// TIA Portal V20 export
FUNCTION_BLOCK "PR_HIPOTTestSeq_Soft2.0 1_workflow_cd2a65"   // FB45, LAD
{ S7_Optimized_Access := 'TRUE' }
// stored: MemoryReserve 100, SetENOAutomatically false
   VAR_INPUT
      iAutoRunning : Bool;
      iFaultReset : Bool;
      iHiPotProbeUp : Bool;
      iHiPotTestOver : Bool;
      iHiPotTestProbeDown : Bool;
      iPartPresent : Bool;
      iPressProbeUp : Bool;
      iReset_fault : Bool;
      iShuttleAtHiPotTest : Bool;
      iSstMode : Bool;
      iSstPB : Bool;
      iStartFrmShuttleSeq : Bool;
      iTestProbeDown : Bool;
      iTestProbeUp : Bool;
      iTestProbesUp : Bool;
      iThicknessTestOver : Bool;
      iScanOK : Bool;
      iScanNOK : Bool;
      iRetryCount : Int;
      iForcedAccept : Bool;
      iRetry : Bool;
   END_VAR
   VAR_OUTPUT
      qHiPotTestOver : Bool;
      qStateNo : Int;
      qMessage : Array[0..2] of Bool;
   END_VAR
   VAR
      c20_ChkRecoveryStatus_T1 : Bool;
      c20_ChkRecoveryStatus_T2 : Bool;
      c20_ChkRecoveryStatus_T3 : Bool;
      c20_ChkRecoveryStatus_T4 : Bool;
      c50_ChkPartPresentShuttlePos_T1 : Bool;
      c50_ChkPartPresentShuttlePos_T2 : Bool;
      s100_WtHiPotTestProbesDown : Bool;
      s100_WtHiPotTestProbesDown_T1 : Bool;
      s10_WtStartFrmShuttleSeq : Bool;
      s10_WtStartFrmShuttleSeq_T1 : Bool;
      s110_WtHiPotTestOver : Bool;
      s110_WtHiPotTestOver_T1 : Bool;
      s120_WtHiPotProbeUp : Bool;
      s120_WtHiPotProbeUp_T1 : Bool;
      s130_WtPressProbesUp : Bool;
      s130_WtPressProbesUp_T1 : Bool;
      s140_WtStartLow : Bool;
      s140_WtStartLow_T1 : Bool;
      s1_WtResetRel : Bool;
      s1_WtResetRel_T1 : Bool;
      s20_ChkRecoveryStatus : Bool;
      s20_ChkRecoveryStatus_T1 : Bool;
      s20_ChkRecoveryStatus_T2 : Bool;
      s20_ChkRecoveryStatus_T3 : Bool;
      s20_ChkRecoveryStatus_T4 : Bool;
      s30_WtOperatorAck : Bool;
      s30_WtOperatorAck_T1 : Bool;
      s40_WtAllSlidesHome : Bool;
      s40_WtAllSlidesHome_T1 : Bool;
      s50_ChkPartPresentShuttlePos : Bool;
      s50_ChkPartPresentShuttlePos_T1 : Bool;
      s50_ChkPartPresentShuttlePos_T2 : Bool;
      s75_WtScanOver : Bool;
      s75_WtScanOver_T1 : Bool;
      s75_WtScanOver_T2 : Bool;
      s76_ChkReryCountOver : Bool;
      s76_ChkRetryCountOver_T1 : Bool;
      s76_ChkRetryCountOver_T2 : Bool;
      s77_WtOperatorDecision : Bool;
      s77_WtOperatorDecision_T1 : Bool;
      s77_WtOperatorDecision_T2 : Bool;
      s70_WtPartPresentShuttlePos : Bool;
      s70_WtPartPresentShuttlePos_T1 : Bool;
      s80_WtTestProbeDown : Bool;
      s80_WtTestProbeDown_T1 : Bool;
      s90_WtThicknessTestOver : Bool;
      s90_WtThicknessTestOver_T1 : Bool;
      sAbnormalStatus : Bool;
      sHiPotTestInProgress : Bool;
      sSst : Bool;
      sSstPulse : Bool;
      sSstRise : Bool;
      sStWtResetRel : Bool;
      sStWtResetRel_T1 : Bool;
      sThicknessTestInProgress : Bool;
      sScanRetryCount : Int;
   END_VAR
   VAR_TEMP
      tOne : Bool;
   END_VAR
   VAR_TEMP   // added for the SCL form of the ladder/FBD networks
      _w1 : Bool;
      _w2 : Bool;
      _w3 : Bool;
   END_VAR
BEGIN

REGION Network 1
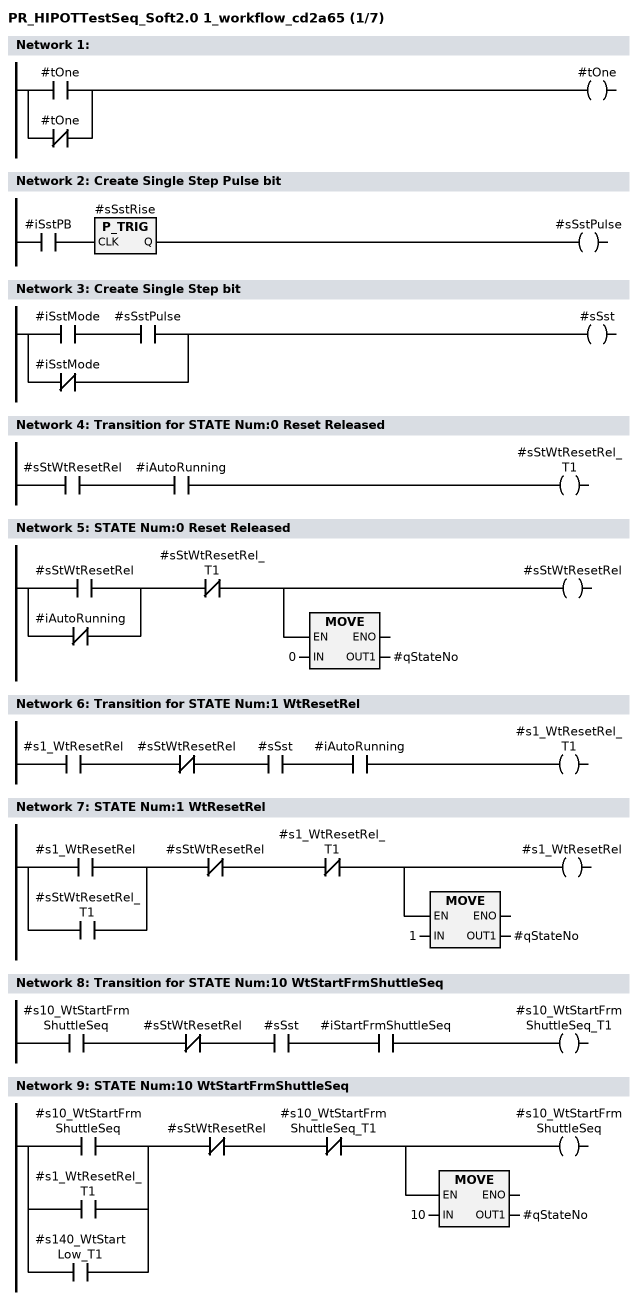
   RUNG wire#powerrail
      Contact( #tOne )
      wire#w1
      Coil( #tOne )
   END_RUNG
   RUNG wire#powerrail
      I_Contact( #tOne )
   END_RUNG wire#w1
   // the same network as SCL:
   #tOne := #tOne OR NOT #tOne;
END_REGION

REGION Network 2: Create Single Step Pulse bit
   RUNG wire#powerrail
      Contact( #iSstPB )
      P_Trig( #sSstRise )
      Coil( #sSstPulse )
   END_RUNG
   // the same network as SCL:
   #_w1 := #iSstPB AND NOT #sSstRise;   // rising edge
   #sSstRise := #iSstPB;
   #sSstPulse := #_w1;
END_REGION

REGION Network 3: Create Single Step bit
   RUNG wire#powerrail
      Contact( #iSstMode )
      Contact( #sSstPulse )
      wire#w1
      Coil( #sSst )
   END_RUNG
   RUNG wire#powerrail
      I_Contact( #iSstMode )
   END_RUNG wire#w1
   // the same network as SCL:
   #sSst := (#iSstMode AND #sSstPulse) OR NOT #iSstMode;
END_REGION

REGION Network 4: Transition for STATE Num:0 Reset Released
   RUNG wire#powerrail
      Contact( #sStWtResetRel )
      Contact( #iAutoRunning )
      Coil( #sStWtResetRel_T1 )
   END_RUNG
   // the same network as SCL:
   #sStWtResetRel_T1 := #sStWtResetRel AND #iAutoRunning;
END_REGION

REGION Network 5: STATE Num:0 Reset Released
   RUNG wire#powerrail
      Contact( #sStWtResetRel )
      wire#w1
      I_Contact( #sStWtResetRel_T1 )
      wire#w2
      Coil( #sStWtResetRel )
   END_RUNG
   RUNG wire#powerrail
      I_Contact( #iAutoRunning )
   END_RUNG wire#w1
   RUNG wire#w2
      { S7_GenerateENO := "TRUE" } Move(in := 0, out1 => #qStateNo)
   END_RUNG
   // the same network as SCL:
   #sStWtResetRel := (#sStWtResetRel OR NOT #iAutoRunning) AND NOT #sStWtResetRel_T1;
   IF #sStWtResetRel THEN #qStateNo := 0; END_IF;
END_REGION

REGION Network 6: Transition for STATE Num:1 WtResetRel
   RUNG wire#powerrail
      Contact( #s1_WtResetRel )
      I_Contact( #sStWtResetRel )
      Contact( #sSst )
      Contact( #iAutoRunning )
      Coil( #s1_WtResetRel_T1 )
   END_RUNG
   // the same network as SCL:
   #s1_WtResetRel_T1 := #s1_WtResetRel AND NOT #sStWtResetRel AND #sSst AND #iAutoRunning;
END_REGION

REGION Network 7: STATE Num:1 WtResetRel
   RUNG wire#powerrail
      Contact( #s1_WtResetRel )
      wire#w1
      I_Contact( #sStWtResetRel )
      I_Contact( #s1_WtResetRel_T1 )
      wire#w2
      Coil( #s1_WtResetRel )
   END_RUNG
   RUNG wire#powerrail
      Contact( #sStWtResetRel_T1 )
   END_RUNG wire#w1
   RUNG wire#w2
      { S7_GenerateENO := "TRUE" } Move(in := 1, out1 => #qStateNo)
   END_RUNG
   // the same network as SCL:
   #s1_WtResetRel := (#s1_WtResetRel OR #sStWtResetRel_T1) AND NOT #sStWtResetRel AND NOT #s1_WtResetRel_T1;
   IF #s1_WtResetRel THEN #qStateNo := 1; END_IF;
END_REGION

REGION Network 8: Transition for STATE Num:10 WtStartFrmShuttleSeq
   RUNG wire#powerrail
      Contact( #s10_WtStartFrmShuttleSeq )
      I_Contact( #sStWtResetRel )
      Contact( #sSst )
      Contact( #iStartFrmShuttleSeq )
      Coil( #s10_WtStartFrmShuttleSeq_T1 )
   END_RUNG
   // the same network as SCL:
   #s10_WtStartFrmShuttleSeq_T1 := #s10_WtStartFrmShuttleSeq AND NOT #sStWtResetRel AND #sSst AND #iStartFrmShuttleSeq;
END_REGION

REGION Network 9: STATE Num:10 WtStartFrmShuttleSeq
   RUNG wire#powerrail
      Contact( #s10_WtStartFrmShuttleSeq )
      wire#w1
      I_Contact( #sStWtResetRel )
      I_Contact( #s10_WtStartFrmShuttleSeq_T1 )
      wire#w2
      Coil( #s10_WtStartFrmShuttleSeq )
   END_RUNG
   RUNG wire#powerrail
      Contact( #s1_WtResetRel_T1 )
   END_RUNG wire#w1
   RUNG wire#powerrail
      Contact( #s140_WtStartLow_T1 )
   END_RUNG wire#w1
   RUNG wire#w2
      { S7_GenerateENO := "TRUE" } Move(in := 10, out1 => #qStateNo)
   END_RUNG
   // the same network as SCL:
   #s10_WtStartFrmShuttleSeq := (#s10_WtStartFrmShuttleSeq OR #s1_WtResetRel_T1 OR #s140_WtStartLow_T1) AND NOT #sStWtResetRel AND NOT #s10_WtStartFrmShuttleSeq_T1;
   IF #s10_WtStartFrmShuttleSeq THEN #qStateNo := 10; END_IF;
END_REGION

REGION Network 10: Condition1 for STATE Num:20 ChkRecoveryStatus
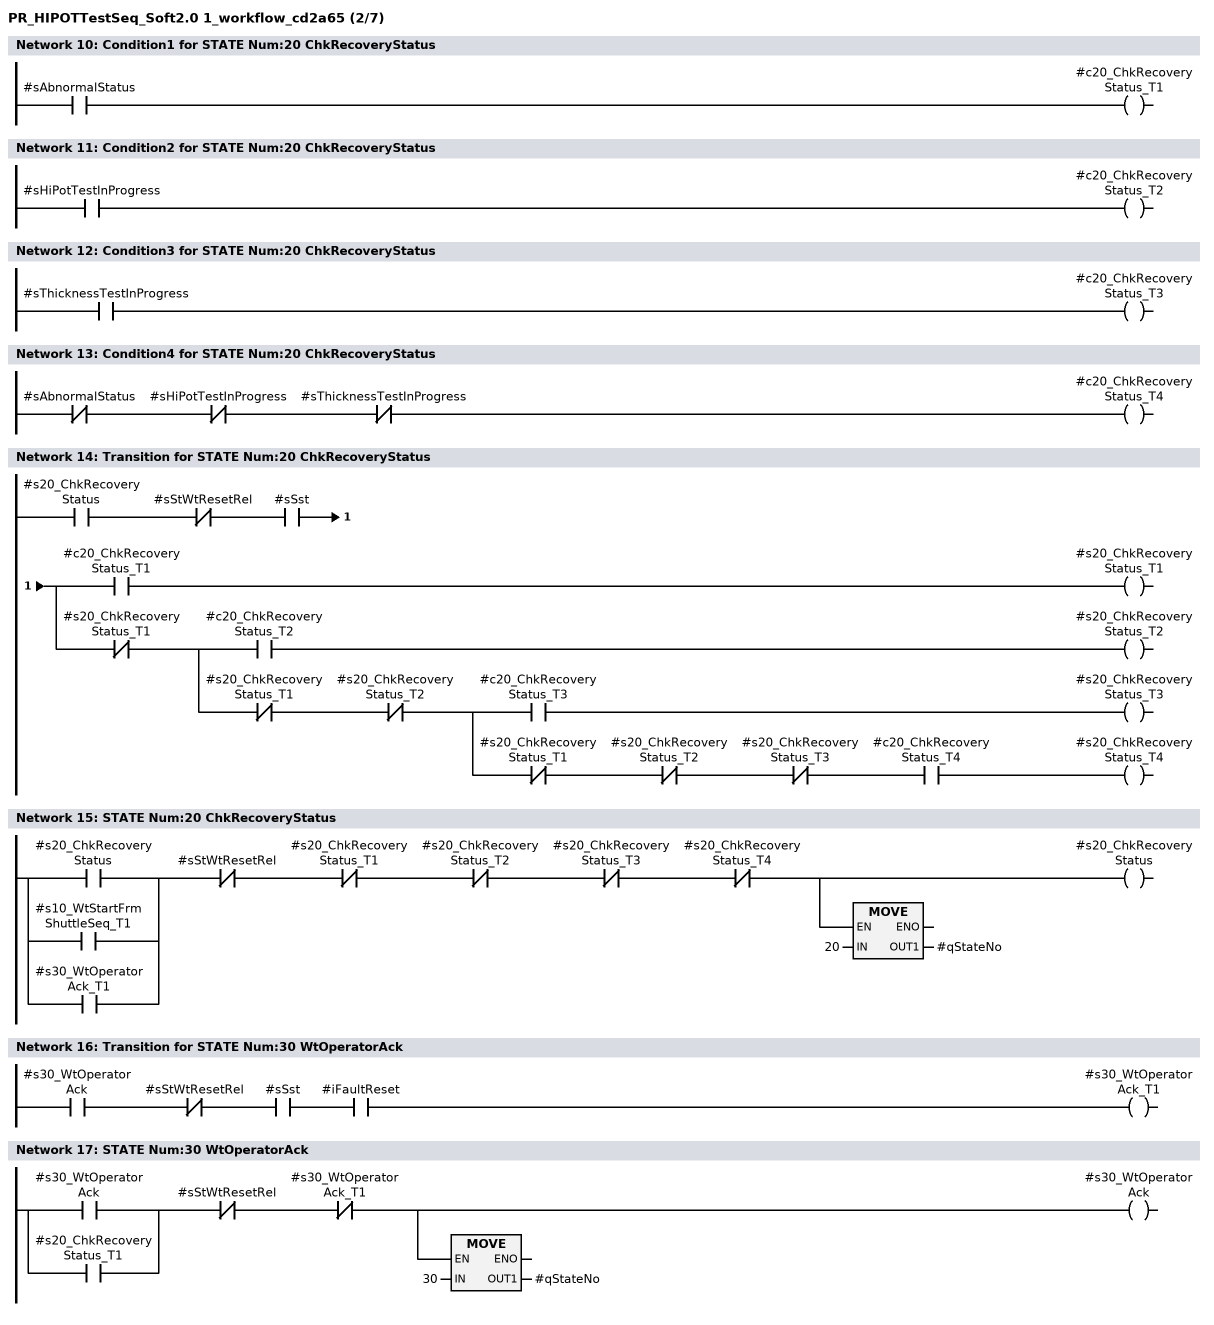
   RUNG wire#powerrail
      Contact( #sAbnormalStatus )
      Coil( #c20_ChkRecoveryStatus_T1 )
   END_RUNG
   // the same network as SCL:
   #c20_ChkRecoveryStatus_T1 := #sAbnormalStatus;
END_REGION

REGION Network 11: Condition2 for STATE Num:20 ChkRecoveryStatus
   RUNG wire#powerrail
      Contact( #sHiPotTestInProgress )
      Coil( #c20_ChkRecoveryStatus_T2 )
   END_RUNG
   // the same network as SCL:
   #c20_ChkRecoveryStatus_T2 := #sHiPotTestInProgress;
END_REGION

REGION Network 12: Condition3 for STATE Num:20 ChkRecoveryStatus
   RUNG wire#powerrail
      Contact( #sThicknessTestInProgress )
      Coil( #c20_ChkRecoveryStatus_T3 )
   END_RUNG
   // the same network as SCL:
   #c20_ChkRecoveryStatus_T3 := #sThicknessTestInProgress;
END_REGION

REGION Network 13: Condition4 for STATE Num:20 ChkRecoveryStatus
   RUNG wire#powerrail
      I_Contact( #sAbnormalStatus )
      I_Contact( #sHiPotTestInProgress )
      I_Contact( #sThicknessTestInProgress )
      Coil( #c20_ChkRecoveryStatus_T4 )
   END_RUNG
   // the same network as SCL:
   #c20_ChkRecoveryStatus_T4 := NOT #sAbnormalStatus AND NOT #sHiPotTestInProgress AND NOT #sThicknessTestInProgress;
END_REGION

REGION Network 14: Transition for STATE Num:20 ChkRecoveryStatus
   RUNG wire#powerrail
      Contact( #s20_ChkRecoveryStatus )
      I_Contact( #sStWtResetRel )
      Contact( #sSst )
      wire#w1
      Contact( #c20_ChkRecoveryStatus_T1 )
      Coil( #s20_ChkRecoveryStatus_T1 )
   END_RUNG
   RUNG wire#w1
      I_Contact( #s20_ChkRecoveryStatus_T1 )
      wire#w2
      Contact( #c20_ChkRecoveryStatus_T2 )
      Coil( #s20_ChkRecoveryStatus_T2 )
   END_RUNG
   RUNG wire#w2
      I_Contact( #s20_ChkRecoveryStatus_T1 )
      I_Contact( #s20_ChkRecoveryStatus_T2 )
      wire#w3
      Contact( #c20_ChkRecoveryStatus_T3 )
      Coil( #s20_ChkRecoveryStatus_T3 )
   END_RUNG
   RUNG wire#w3
      I_Contact( #s20_ChkRecoveryStatus_T1 )
      I_Contact( #s20_ChkRecoveryStatus_T2 )
      I_Contact( #s20_ChkRecoveryStatus_T3 )
      Contact( #c20_ChkRecoveryStatus_T4 )
      Coil( #s20_ChkRecoveryStatus_T4 )
   END_RUNG
   // the same network as SCL:
   #_w1 := #s20_ChkRecoveryStatus AND NOT #sStWtResetRel AND #sSst;
   #s20_ChkRecoveryStatus_T1 := #_w1 AND #c20_ChkRecoveryStatus_T1;
   #_w2 := #_w1 AND NOT #s20_ChkRecoveryStatus_T1;
   #s20_ChkRecoveryStatus_T2 := #_w2 AND #c20_ChkRecoveryStatus_T2;
   #_w3 := #_w2 AND NOT #s20_ChkRecoveryStatus_T1 AND NOT #s20_ChkRecoveryStatus_T2;
   #s20_ChkRecoveryStatus_T3 := #_w3 AND #c20_ChkRecoveryStatus_T3;
   #s20_ChkRecoveryStatus_T4 := #_w3 AND NOT #s20_ChkRecoveryStatus_T1 AND NOT #s20_ChkRecoveryStatus_T2 AND NOT #s20_ChkRecoveryStatus_T3 AND #c20_ChkRecoveryStatus_T4;
END_REGION

REGION Network 15: STATE Num:20 ChkRecoveryStatus
   RUNG wire#powerrail
      Contact( #s20_ChkRecoveryStatus )
      wire#w1
      I_Contact( #sStWtResetRel )
      I_Contact( #s20_ChkRecoveryStatus_T1 )
      I_Contact( #s20_ChkRecoveryStatus_T2 )
      I_Contact( #s20_ChkRecoveryStatus_T3 )
      I_Contact( #s20_ChkRecoveryStatus_T4 )
      wire#w2
      Coil( #s20_ChkRecoveryStatus )
   END_RUNG
   RUNG wire#powerrail
      Contact( #s10_WtStartFrmShuttleSeq_T1 )
   END_RUNG wire#w1
   RUNG wire#powerrail
      Contact( #s30_WtOperatorAck_T1 )
   END_RUNG wire#w1
   RUNG wire#w2
      { S7_GenerateENO := "TRUE" } Move(in := 20, out1 => #qStateNo)
   END_RUNG
   // the same network as SCL:
   #s20_ChkRecoveryStatus := (#s20_ChkRecoveryStatus OR #s10_WtStartFrmShuttleSeq_T1 OR #s30_WtOperatorAck_T1) AND NOT #sStWtResetRel AND NOT #s20_ChkRecoveryStatus_T1 AND NOT #s20_ChkRecoveryStatus_T2 AND NOT #s20_ChkRecoveryStatus_T3 AND NOT #s20_ChkRecoveryStatus_T4;
   IF #s20_ChkRecoveryStatus THEN #qStateNo := 20; END_IF;
END_REGION

REGION Network 16: Transition for STATE Num:30 WtOperatorAck
   RUNG wire#powerrail
      Contact( #s30_WtOperatorAck )
      I_Contact( #sStWtResetRel )
      Contact( #sSst )
      Contact( #iFaultReset )
      Coil( #s30_WtOperatorAck_T1 )
   END_RUNG
   // the same network as SCL:
   #s30_WtOperatorAck_T1 := #s30_WtOperatorAck AND NOT #sStWtResetRel AND #sSst AND #iFaultReset;
END_REGION

REGION Network 17: STATE Num:30 WtOperatorAck
   RUNG wire#powerrail
      Contact( #s30_WtOperatorAck )
      wire#w1
      I_Contact( #sStWtResetRel )
      I_Contact( #s30_WtOperatorAck_T1 )
      wire#w2
      Coil( #s30_WtOperatorAck )
   END_RUNG
   RUNG wire#powerrail
      Contact( #s20_ChkRecoveryStatus_T1 )
   END_RUNG wire#w1
   RUNG wire#w2
      { S7_GenerateENO := "TRUE" } Move(in := 30, out1 => #qStateNo)
   END_RUNG
   // the same network as SCL:
   #s30_WtOperatorAck := (#s30_WtOperatorAck OR #s20_ChkRecoveryStatus_T1) AND NOT #sStWtResetRel AND NOT #s30_WtOperatorAck_T1;
   IF #s30_WtOperatorAck THEN #qStateNo := 30; END_IF;
END_REGION

REGION Network 18: Transition for STATE Num:40 WtAllSlidesHome
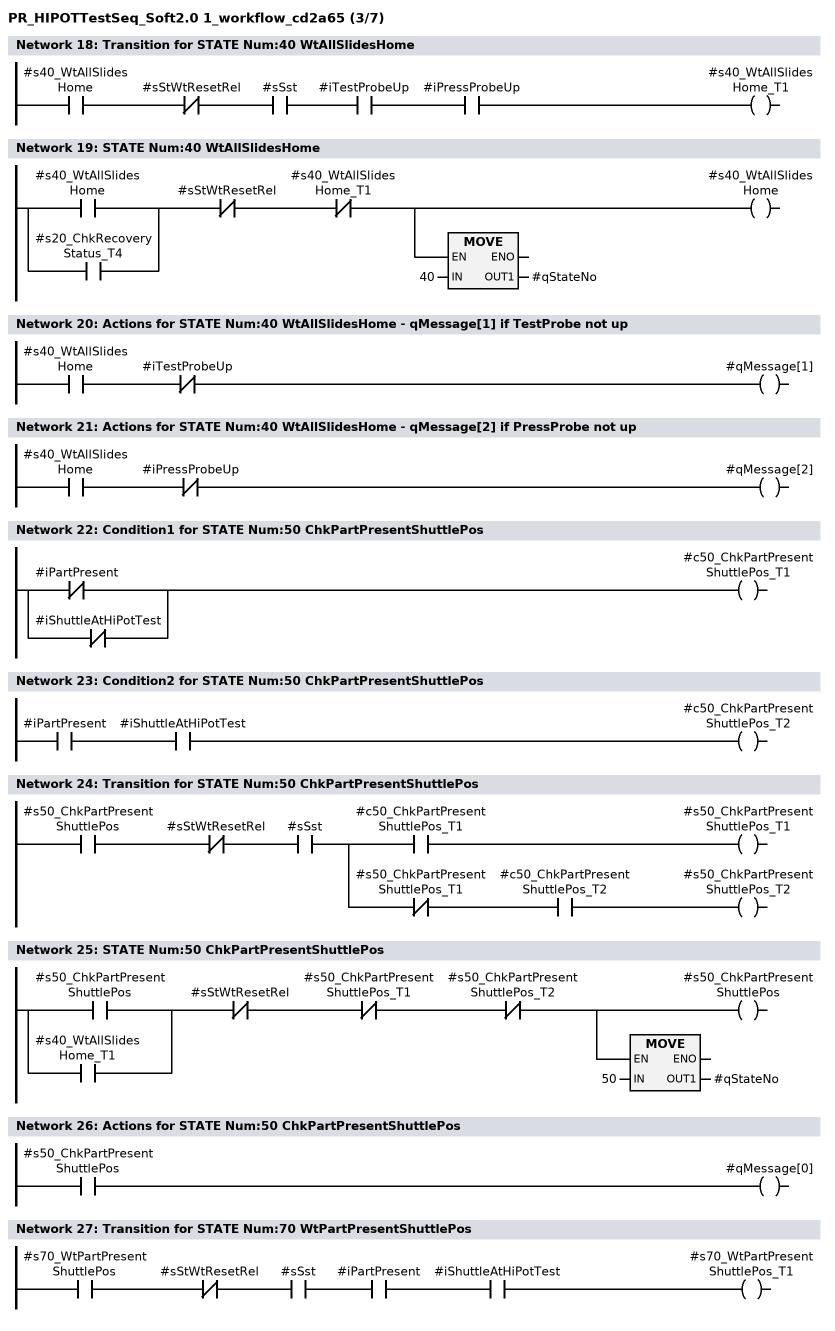
   RUNG wire#powerrail
      Contact( #s40_WtAllSlidesHome )
      I_Contact( #sStWtResetRel )
      Contact( #sSst )
      Contact( #iTestProbeUp )
      Contact( #iPressProbeUp )
      Coil( #s40_WtAllSlidesHome_T1 )
   END_RUNG
   // the same network as SCL:
   #s40_WtAllSlidesHome_T1 := #s40_WtAllSlidesHome AND NOT #sStWtResetRel AND #sSst AND #iTestProbeUp AND #iPressProbeUp;
END_REGION

REGION Network 19: STATE Num:40 WtAllSlidesHome
   RUNG wire#powerrail
      Contact( #s40_WtAllSlidesHome )
      wire#w1
      I_Contact( #sStWtResetRel )
      I_Contact( #s40_WtAllSlidesHome_T1 )
      wire#w2
      Coil( #s40_WtAllSlidesHome )
   END_RUNG
   RUNG wire#powerrail
      Contact( #s20_ChkRecoveryStatus_T4 )
   END_RUNG wire#w1
   RUNG wire#w2
      { S7_GenerateENO := "TRUE" } Move(in := 40, out1 => #qStateNo)
   END_RUNG
   // the same network as SCL:
   #s40_WtAllSlidesHome := (#s40_WtAllSlidesHome OR #s20_ChkRecoveryStatus_T4) AND NOT #sStWtResetRel AND NOT #s40_WtAllSlidesHome_T1;
   IF #s40_WtAllSlidesHome THEN #qStateNo := 40; END_IF;
END_REGION

REGION Network 20: Actions for STATE Num:40 WtAllSlidesHome - qMessage[1] if TestProbe not up
   RUNG wire#powerrail
      Contact( #s40_WtAllSlidesHome )
      I_Contact( #iTestProbeUp )
      Coil( #qMessage[1] )
   END_RUNG
   // the same network as SCL:
   #qMessage[1] := #s40_WtAllSlidesHome AND NOT #iTestProbeUp;
END_REGION

REGION Network 21: Actions for STATE Num:40 WtAllSlidesHome - qMessage[2] if PressProbe not up
   RUNG wire#powerrail
      Contact( #s40_WtAllSlidesHome )
      I_Contact( #iPressProbeUp )
      Coil( #qMessage[2] )
   END_RUNG
   // the same network as SCL:
   #qMessage[2] := #s40_WtAllSlidesHome AND NOT #iPressProbeUp;
END_REGION

REGION Network 22: Condition1 for STATE Num:50 ChkPartPresentShuttlePos
   RUNG wire#powerrail
      I_Contact( #iPartPresent )
      wire#w1
      Coil( #c50_ChkPartPresentShuttlePos_T1 )
   END_RUNG
   RUNG wire#powerrail
      I_Contact( #iShuttleAtHiPotTest )
   END_RUNG wire#w1
   // the same network as SCL:
   #c50_ChkPartPresentShuttlePos_T1 := NOT #iPartPresent OR NOT #iShuttleAtHiPotTest;
END_REGION

REGION Network 23: Condition2 for STATE Num:50 ChkPartPresentShuttlePos
   RUNG wire#powerrail
      Contact( #iPartPresent )
      Contact( #iShuttleAtHiPotTest )
      Coil( #c50_ChkPartPresentShuttlePos_T2 )
   END_RUNG
   // the same network as SCL:
   #c50_ChkPartPresentShuttlePos_T2 := #iPartPresent AND #iShuttleAtHiPotTest;
END_REGION

REGION Network 24: Transition for STATE Num:50 ChkPartPresentShuttlePos
   RUNG wire#powerrail
      Contact( #s50_ChkPartPresentShuttlePos )
      I_Contact( #sStWtResetRel )
      Contact( #sSst )
      wire#w1
      Contact( #c50_ChkPartPresentShuttlePos_T1 )
      Coil( #s50_ChkPartPresentShuttlePos_T1 )
   END_RUNG
   RUNG wire#w1
      I_Contact( #s50_ChkPartPresentShuttlePos_T1 )
      Contact( #c50_ChkPartPresentShuttlePos_T2 )
      Coil( #s50_ChkPartPresentShuttlePos_T2 )
   END_RUNG
   // the same network as SCL:
   #_w1 := #s50_ChkPartPresentShuttlePos AND NOT #sStWtResetRel AND #sSst;
   #s50_ChkPartPresentShuttlePos_T1 := #_w1 AND #c50_ChkPartPresentShuttlePos_T1;
   #s50_ChkPartPresentShuttlePos_T2 := #_w1 AND NOT #s50_ChkPartPresentShuttlePos_T1 AND #c50_ChkPartPresentShuttlePos_T2;
END_REGION

REGION Network 25: STATE Num:50 ChkPartPresentShuttlePos
   RUNG wire#powerrail
      Contact( #s50_ChkPartPresentShuttlePos )
      wire#w1
      I_Contact( #sStWtResetRel )
      I_Contact( #s50_ChkPartPresentShuttlePos_T1 )
      I_Contact( #s50_ChkPartPresentShuttlePos_T2 )
      wire#w2
      Coil( #s50_ChkPartPresentShuttlePos )
   END_RUNG
   RUNG wire#powerrail
      Contact( #s40_WtAllSlidesHome_T1 )
   END_RUNG wire#w1
   RUNG wire#w2
      { S7_GenerateENO := "TRUE" } Move(in := 50, out1 => #qStateNo)
   END_RUNG
   // the same network as SCL:
   #s50_ChkPartPresentShuttlePos := (#s50_ChkPartPresentShuttlePos OR #s40_WtAllSlidesHome_T1) AND NOT #sStWtResetRel AND NOT #s50_ChkPartPresentShuttlePos_T1 AND NOT #s50_ChkPartPresentShuttlePos_T2;
   IF #s50_ChkPartPresentShuttlePos THEN #qStateNo := 50; END_IF;
END_REGION

REGION Network 26: Actions for STATE Num:50 ChkPartPresentShuttlePos
   RUNG wire#powerrail
      Contact( #s50_ChkPartPresentShuttlePos )
      Coil( #qMessage[0] )
   END_RUNG
   // the same network as SCL:
   #qMessage[0] := #s50_ChkPartPresentShuttlePos;
END_REGION

REGION Network 27: Transition for STATE Num:70 WtPartPresentShuttlePos
   RUNG wire#powerrail
      Contact( #s70_WtPartPresentShuttlePos )
      I_Contact( #sStWtResetRel )
      Contact( #sSst )
      Contact( #iPartPresent )
      Contact( #iShuttleAtHiPotTest )
      Coil( #s70_WtPartPresentShuttlePos_T1 )
   END_RUNG
   // the same network as SCL:
   #s70_WtPartPresentShuttlePos_T1 := #s70_WtPartPresentShuttlePos AND NOT #sStWtResetRel AND #sSst AND #iPartPresent AND #iShuttleAtHiPotTest;
END_REGION

REGION Network 28: STATE Num:70 WtPartPresentShuttlePos
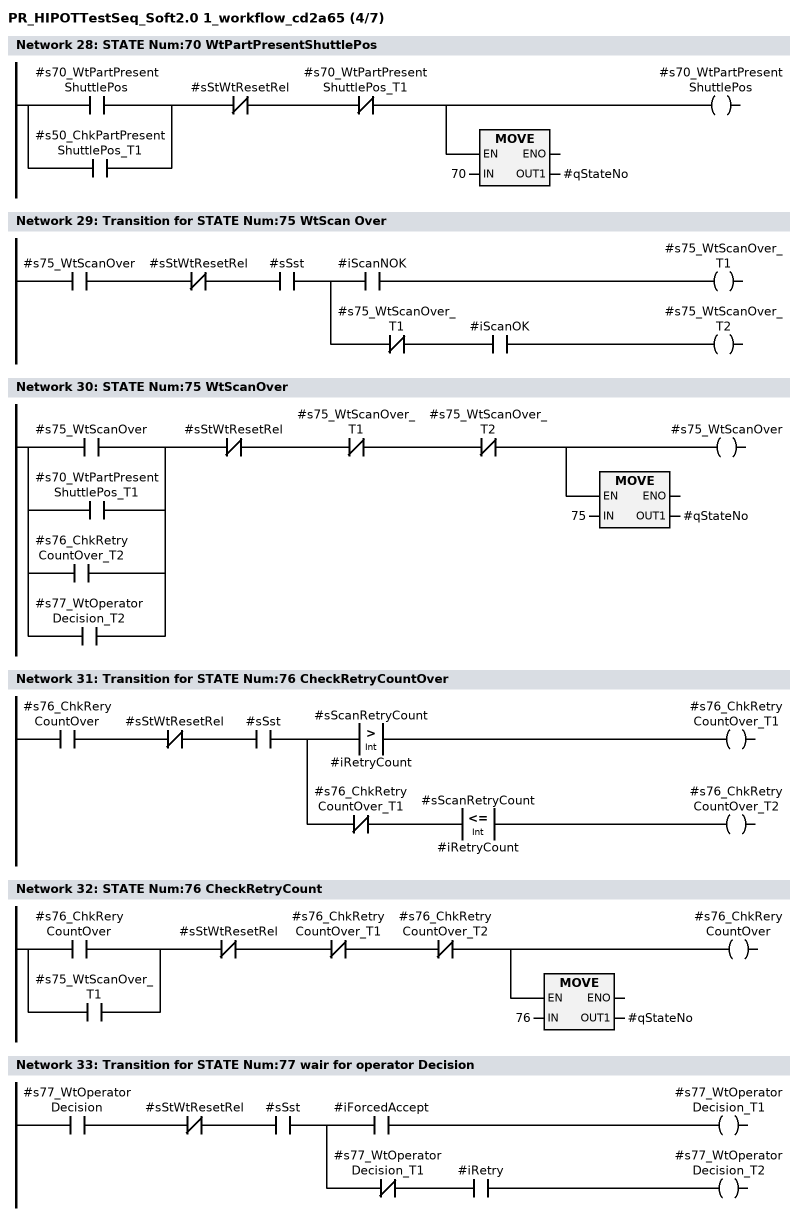
   RUNG wire#powerrail
      Contact( #s70_WtPartPresentShuttlePos )
      wire#w1
      I_Contact( #sStWtResetRel )
      I_Contact( #s70_WtPartPresentShuttlePos_T1 )
      wire#w2
      Coil( #s70_WtPartPresentShuttlePos )
   END_RUNG
   RUNG wire#powerrail
      Contact( #s50_ChkPartPresentShuttlePos_T1 )
   END_RUNG wire#w1
   RUNG wire#w2
      { S7_GenerateENO := "TRUE" } Move(in := 70, out1 => #qStateNo)
   END_RUNG
   // the same network as SCL:
   #s70_WtPartPresentShuttlePos := (#s70_WtPartPresentShuttlePos OR #s50_ChkPartPresentShuttlePos_T1) AND NOT #sStWtResetRel AND NOT #s70_WtPartPresentShuttlePos_T1;
   IF #s70_WtPartPresentShuttlePos THEN #qStateNo := 70; END_IF;
END_REGION

REGION Network 29: Transition for STATE Num:75 WtScan Over
   RUNG wire#powerrail
      Contact( #s75_WtScanOver )
      I_Contact( #sStWtResetRel )
      Contact( #sSst )
      wire#w1
      Contact( #iScanNOK )
      Coil( #s75_WtScanOver_T1 )
   END_RUNG
   RUNG wire#w1
      I_Contact( #s75_WtScanOver_T1 )
      Contact( #iScanOK )
      Coil( #s75_WtScanOver_T2 )
   END_RUNG
   // the same network as SCL:
   #_w1 := #s75_WtScanOver AND NOT #sStWtResetRel AND #sSst;
   #s75_WtScanOver_T1 := #_w1 AND #iScanNOK;
   #s75_WtScanOver_T2 := #_w1 AND NOT #s75_WtScanOver_T1 AND #iScanOK;
END_REGION

REGION Network 30: STATE Num:75 WtScanOver
   RUNG wire#powerrail
      Contact( #s75_WtScanOver )
      wire#w1
      I_Contact( #sStWtResetRel )
      I_Contact( #s75_WtScanOver_T1 )
      I_Contact( #s75_WtScanOver_T2 )
      wire#w2
      Coil( #s75_WtScanOver )
   END_RUNG
   RUNG wire#powerrail
      Contact( #s70_WtPartPresentShuttlePos_T1 )
   END_RUNG wire#w1
   RUNG wire#powerrail
      Contact( #s76_ChkRetryCountOver_T2 )
   END_RUNG wire#w1
   RUNG wire#powerrail
      Contact( #s77_WtOperatorDecision_T2 )
   END_RUNG wire#w1
   RUNG wire#w2
      Move(in := 75, out1 => #qStateNo)
   END_RUNG
   // the same network as SCL:
   #s75_WtScanOver := (#s75_WtScanOver OR #s70_WtPartPresentShuttlePos_T1 OR #s76_ChkRetryCountOver_T2 OR #s77_WtOperatorDecision_T2) AND NOT #sStWtResetRel AND NOT #s75_WtScanOver_T1 AND NOT #s75_WtScanOver_T2;
   IF #s75_WtScanOver THEN #qStateNo := 75; END_IF;
END_REGION

REGION Network 31: Transition for STATE Num:76 CheckRetryCountOver
   RUNG wire#powerrail
      Contact( #s76_ChkReryCountOver )
      I_Contact( #sStWtResetRel )
      Contact( #sSst )
      wire#w1
      { S7_Templates := "SrcType := Int" } GT_Contact(in1 := #sScanRetryCount, in2 := #iRetryCount)
      Coil( #s76_ChkRetryCountOver_T1 )
   END_RUNG
   RUNG wire#w1
      I_Contact( #s76_ChkRetryCountOver_T1 )
      { S7_Templates := "SrcType := Int" } LE_Contact(in1 := #sScanRetryCount, in2 := #iRetryCount)
      Coil( #s76_ChkRetryCountOver_T2 )
   END_RUNG
   // the same network as SCL:
   #_w1 := #s76_ChkReryCountOver AND NOT #sStWtResetRel AND #sSst;
   #s76_ChkRetryCountOver_T1 := #_w1 AND (#sScanRetryCount > #iRetryCount);
   #s76_ChkRetryCountOver_T2 := #_w1 AND NOT #s76_ChkRetryCountOver_T1 AND (#sScanRetryCount <= #iRetryCount);
END_REGION

REGION Network 32: STATE Num:76 CheckRetryCount
   RUNG wire#powerrail
      Contact( #s76_ChkReryCountOver )
      wire#w1
      I_Contact( #sStWtResetRel )
      I_Contact( #s76_ChkRetryCountOver_T1 )
      I_Contact( #s76_ChkRetryCountOver_T2 )
      wire#w2
      Coil( #s76_ChkReryCountOver )
   END_RUNG
   RUNG wire#powerrail
      Contact( #s75_WtScanOver_T1 )
   END_RUNG wire#w1
   RUNG wire#w2
      Move(in := 76, out1 => #qStateNo)
   END_RUNG
   // the same network as SCL:
   #s76_ChkReryCountOver := (#s76_ChkReryCountOver OR #s75_WtScanOver_T1) AND NOT #sStWtResetRel AND NOT #s76_ChkRetryCountOver_T1 AND NOT #s76_ChkRetryCountOver_T2;
   IF #s76_ChkReryCountOver THEN #qStateNo := 76; END_IF;
END_REGION

REGION Network 33: Transition for STATE Num:77 wair for operator Decision
   RUNG wire#powerrail
      Contact( #s77_WtOperatorDecision )
      I_Contact( #sStWtResetRel )
      Contact( #sSst )
      wire#w1
      Contact( #iForcedAccept )
      Coil( #s77_WtOperatorDecision_T1 )
   END_RUNG
   RUNG wire#w1
      I_Contact( #s77_WtOperatorDecision_T1 )
      Contact( #iRetry )
      Coil( #s77_WtOperatorDecision_T2 )
   END_RUNG
   // the same network as SCL:
   #_w1 := #s77_WtOperatorDecision AND NOT #sStWtResetRel AND #sSst;
   #s77_WtOperatorDecision_T1 := #_w1 AND #iForcedAccept;
   #s77_WtOperatorDecision_T2 := #_w1 AND NOT #s77_WtOperatorDecision_T1 AND #iRetry;
END_REGION

REGION Network 34: STATE Num:77 wait For Operator Decision
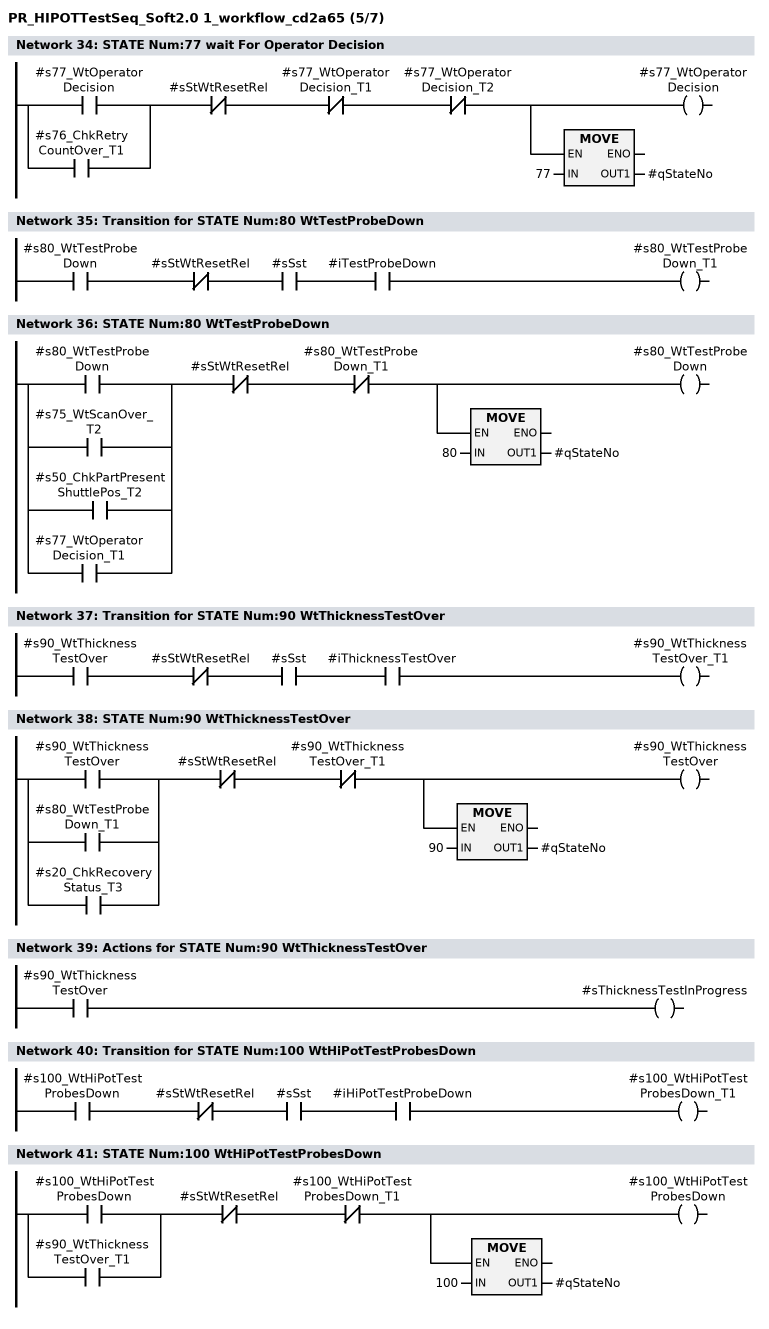
   RUNG wire#powerrail
      Contact( #s77_WtOperatorDecision )
      wire#w1
      I_Contact( #sStWtResetRel )
      I_Contact( #s77_WtOperatorDecision_T1 )
      I_Contact( #s77_WtOperatorDecision_T2 )
      wire#w2
      Coil( #s77_WtOperatorDecision )
   END_RUNG
   RUNG wire#powerrail
      Contact( #s76_ChkRetryCountOver_T1 )
   END_RUNG wire#w1
   RUNG wire#w2
      Move(in := 77, out1 => #qStateNo)
   END_RUNG
   // the same network as SCL:
   #s77_WtOperatorDecision := (#s77_WtOperatorDecision OR #s76_ChkRetryCountOver_T1) AND NOT #sStWtResetRel AND NOT #s77_WtOperatorDecision_T1 AND NOT #s77_WtOperatorDecision_T2;
   IF #s77_WtOperatorDecision THEN #qStateNo := 77; END_IF;
END_REGION

REGION Network 35: Transition for STATE Num:80 WtTestProbeDown
   RUNG wire#powerrail
      Contact( #s80_WtTestProbeDown )
      I_Contact( #sStWtResetRel )
      Contact( #sSst )
      Contact( #iTestProbeDown )
      Coil( #s80_WtTestProbeDown_T1 )
   END_RUNG
   // the same network as SCL:
   #s80_WtTestProbeDown_T1 := #s80_WtTestProbeDown AND NOT #sStWtResetRel AND #sSst AND #iTestProbeDown;
END_REGION

REGION Network 36: STATE Num:80 WtTestProbeDown
   RUNG wire#powerrail
      Contact( #s80_WtTestProbeDown )
      wire#w1
      I_Contact( #sStWtResetRel )
      I_Contact( #s80_WtTestProbeDown_T1 )
      wire#w2
      Coil( #s80_WtTestProbeDown )
   END_RUNG
   RUNG wire#powerrail
      Contact( #s75_WtScanOver_T2 )
   END_RUNG wire#w1
   RUNG wire#powerrail
      Contact( #s50_ChkPartPresentShuttlePos_T2 )
   END_RUNG wire#w1
   RUNG wire#powerrail
      Contact( #s77_WtOperatorDecision_T1 )
   END_RUNG wire#w1
   RUNG wire#w2
      { S7_GenerateENO := "TRUE" } Move(in := 80, out1 => #qStateNo)
   END_RUNG
   // the same network as SCL:
   #s80_WtTestProbeDown := (#s80_WtTestProbeDown OR #s75_WtScanOver_T2 OR #s50_ChkPartPresentShuttlePos_T2 OR #s77_WtOperatorDecision_T1) AND NOT #sStWtResetRel AND NOT #s80_WtTestProbeDown_T1;
   IF #s80_WtTestProbeDown THEN #qStateNo := 80; END_IF;
END_REGION

REGION Network 37: Transition for STATE Num:90 WtThicknessTestOver
   RUNG wire#powerrail
      Contact( #s90_WtThicknessTestOver )
      I_Contact( #sStWtResetRel )
      Contact( #sSst )
      Contact( #iThicknessTestOver )
      Coil( #s90_WtThicknessTestOver_T1 )
   END_RUNG
   // the same network as SCL:
   #s90_WtThicknessTestOver_T1 := #s90_WtThicknessTestOver AND NOT #sStWtResetRel AND #sSst AND #iThicknessTestOver;
END_REGION

REGION Network 38: STATE Num:90 WtThicknessTestOver
   RUNG wire#powerrail
      Contact( #s90_WtThicknessTestOver )
      wire#w1
      I_Contact( #sStWtResetRel )
      I_Contact( #s90_WtThicknessTestOver_T1 )
      wire#w2
      Coil( #s90_WtThicknessTestOver )
   END_RUNG
   RUNG wire#powerrail
      Contact( #s80_WtTestProbeDown_T1 )
   END_RUNG wire#w1
   RUNG wire#powerrail
      Contact( #s20_ChkRecoveryStatus_T3 )
   END_RUNG wire#w1
   RUNG wire#w2
      { S7_GenerateENO := "TRUE" } Move(in := 90, out1 => #qStateNo)
   END_RUNG
   // the same network as SCL:
   #s90_WtThicknessTestOver := (#s90_WtThicknessTestOver OR #s80_WtTestProbeDown_T1 OR #s20_ChkRecoveryStatus_T3) AND NOT #sStWtResetRel AND NOT #s90_WtThicknessTestOver_T1;
   IF #s90_WtThicknessTestOver THEN #qStateNo := 90; END_IF;
END_REGION

REGION Network 39: Actions for STATE Num:90 WtThicknessTestOver
   RUNG wire#powerrail
      Contact( #s90_WtThicknessTestOver )
      Coil( #sThicknessTestInProgress )
   END_RUNG
   // the same network as SCL:
   #sThicknessTestInProgress := #s90_WtThicknessTestOver;
END_REGION

REGION Network 40: Transition for STATE Num:100 WtHiPotTestProbesDown
   RUNG wire#powerrail
      Contact( #s100_WtHiPotTestProbesDown )
      I_Contact( #sStWtResetRel )
      Contact( #sSst )
      Contact( #iHiPotTestProbeDown )
      Coil( #s100_WtHiPotTestProbesDown_T1 )
   END_RUNG
   // the same network as SCL:
   #s100_WtHiPotTestProbesDown_T1 := #s100_WtHiPotTestProbesDown AND NOT #sStWtResetRel AND #sSst AND #iHiPotTestProbeDown;
END_REGION

REGION Network 41: STATE Num:100 WtHiPotTestProbesDown
   RUNG wire#powerrail
      Contact( #s100_WtHiPotTestProbesDown )
      wire#w1
      I_Contact( #sStWtResetRel )
      I_Contact( #s100_WtHiPotTestProbesDown_T1 )
      wire#w2
      Coil( #s100_WtHiPotTestProbesDown )
   END_RUNG
   RUNG wire#powerrail
      Contact( #s90_WtThicknessTestOver_T1 )
   END_RUNG wire#w1
   RUNG wire#w2
      { S7_GenerateENO := "TRUE" } Move(in := 100, out1 => #qStateNo)
   END_RUNG
   // the same network as SCL:
   #s100_WtHiPotTestProbesDown := (#s100_WtHiPotTestProbesDown OR #s90_WtThicknessTestOver_T1) AND NOT #sStWtResetRel AND NOT #s100_WtHiPotTestProbesDown_T1;
   IF #s100_WtHiPotTestProbesDown THEN #qStateNo := 100; END_IF;
END_REGION

REGION Network 42: Transition for STATE Num:110 WtHiPotTestOver
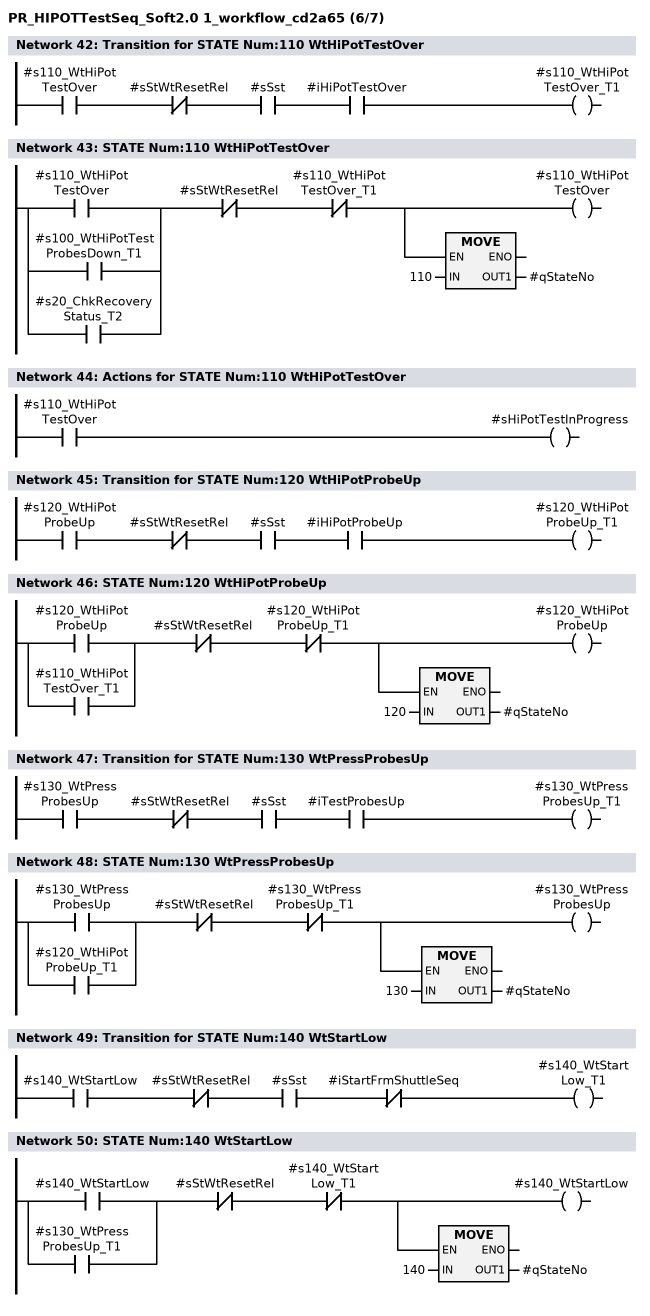
   RUNG wire#powerrail
      Contact( #s110_WtHiPotTestOver )
      I_Contact( #sStWtResetRel )
      Contact( #sSst )
      Contact( #iHiPotTestOver )
      Coil( #s110_WtHiPotTestOver_T1 )
   END_RUNG
   // the same network as SCL:
   #s110_WtHiPotTestOver_T1 := #s110_WtHiPotTestOver AND NOT #sStWtResetRel AND #sSst AND #iHiPotTestOver;
END_REGION

REGION Network 43: STATE Num:110 WtHiPotTestOver
   RUNG wire#powerrail
      Contact( #s110_WtHiPotTestOver )
      wire#w1
      I_Contact( #sStWtResetRel )
      I_Contact( #s110_WtHiPotTestOver_T1 )
      wire#w2
      Coil( #s110_WtHiPotTestOver )
   END_RUNG
   RUNG wire#powerrail
      Contact( #s100_WtHiPotTestProbesDown_T1 )
   END_RUNG wire#w1
   RUNG wire#powerrail
      Contact( #s20_ChkRecoveryStatus_T2 )
   END_RUNG wire#w1
   RUNG wire#w2
      { S7_GenerateENO := "TRUE" } Move(in := 110, out1 => #qStateNo)
   END_RUNG
   // the same network as SCL:
   #s110_WtHiPotTestOver := (#s110_WtHiPotTestOver OR #s100_WtHiPotTestProbesDown_T1 OR #s20_ChkRecoveryStatus_T2) AND NOT #sStWtResetRel AND NOT #s110_WtHiPotTestOver_T1;
   IF #s110_WtHiPotTestOver THEN #qStateNo := 110; END_IF;
END_REGION

REGION Network 44: Actions for STATE Num:110 WtHiPotTestOver
   RUNG wire#powerrail
      Contact( #s110_WtHiPotTestOver )
      Coil( #sHiPotTestInProgress )
   END_RUNG
   // the same network as SCL:
   #sHiPotTestInProgress := #s110_WtHiPotTestOver;
END_REGION

REGION Network 45: Transition for STATE Num:120 WtHiPotProbeUp
   RUNG wire#powerrail
      Contact( #s120_WtHiPotProbeUp )
      I_Contact( #sStWtResetRel )
      Contact( #sSst )
      Contact( #iHiPotProbeUp )
      Coil( #s120_WtHiPotProbeUp_T1 )
   END_RUNG
   // the same network as SCL:
   #s120_WtHiPotProbeUp_T1 := #s120_WtHiPotProbeUp AND NOT #sStWtResetRel AND #sSst AND #iHiPotProbeUp;
END_REGION

REGION Network 46: STATE Num:120 WtHiPotProbeUp
   RUNG wire#powerrail
      Contact( #s120_WtHiPotProbeUp )
      wire#w1
      I_Contact( #sStWtResetRel )
      I_Contact( #s120_WtHiPotProbeUp_T1 )
      wire#w2
      Coil( #s120_WtHiPotProbeUp )
   END_RUNG
   RUNG wire#powerrail
      Contact( #s110_WtHiPotTestOver_T1 )
   END_RUNG wire#w1
   RUNG wire#w2
      { S7_GenerateENO := "TRUE" } Move(in := 120, out1 => #qStateNo)
   END_RUNG
   // the same network as SCL:
   #s120_WtHiPotProbeUp := (#s120_WtHiPotProbeUp OR #s110_WtHiPotTestOver_T1) AND NOT #sStWtResetRel AND NOT #s120_WtHiPotProbeUp_T1;
   IF #s120_WtHiPotProbeUp THEN #qStateNo := 120; END_IF;
END_REGION

REGION Network 47: Transition for STATE Num:130 WtPressProbesUp
   RUNG wire#powerrail
      Contact( #s130_WtPressProbesUp )
      I_Contact( #sStWtResetRel )
      Contact( #sSst )
      Contact( #iTestProbesUp )
      Coil( #s130_WtPressProbesUp_T1 )
   END_RUNG
   // the same network as SCL:
   #s130_WtPressProbesUp_T1 := #s130_WtPressProbesUp AND NOT #sStWtResetRel AND #sSst AND #iTestProbesUp;
END_REGION

REGION Network 48: STATE Num:130 WtPressProbesUp
   RUNG wire#powerrail
      Contact( #s130_WtPressProbesUp )
      wire#w1
      I_Contact( #sStWtResetRel )
      I_Contact( #s130_WtPressProbesUp_T1 )
      wire#w2
      Coil( #s130_WtPressProbesUp )
   END_RUNG
   RUNG wire#powerrail
      Contact( #s120_WtHiPotProbeUp_T1 )
   END_RUNG wire#w1
   RUNG wire#w2
      { S7_GenerateENO := "TRUE" } Move(in := 130, out1 => #qStateNo)
   END_RUNG
   // the same network as SCL:
   #s130_WtPressProbesUp := (#s130_WtPressProbesUp OR #s120_WtHiPotProbeUp_T1) AND NOT #sStWtResetRel AND NOT #s130_WtPressProbesUp_T1;
   IF #s130_WtPressProbesUp THEN #qStateNo := 130; END_IF;
END_REGION

REGION Network 49: Transition for STATE Num:140 WtStartLow
   RUNG wire#powerrail
      Contact( #s140_WtStartLow )
      I_Contact( #sStWtResetRel )
      Contact( #sSst )
      I_Contact( #iStartFrmShuttleSeq )
      Coil( #s140_WtStartLow_T1 )
   END_RUNG
   // the same network as SCL:
   #s140_WtStartLow_T1 := #s140_WtStartLow AND NOT #sStWtResetRel AND #sSst AND NOT #iStartFrmShuttleSeq;
END_REGION

REGION Network 50: STATE Num:140 WtStartLow
   RUNG wire#powerrail
      Contact( #s140_WtStartLow )
      wire#w1
      I_Contact( #sStWtResetRel )
      I_Contact( #s140_WtStartLow_T1 )
      wire#w2
      Coil( #s140_WtStartLow )
   END_RUNG
   RUNG wire#powerrail
      Contact( #s130_WtPressProbesUp_T1 )
   END_RUNG wire#w1
   RUNG wire#w2
      { S7_GenerateENO := "TRUE" } Move(in := 140, out1 => #qStateNo)
   END_RUNG
   // the same network as SCL:
   #s140_WtStartLow := (#s140_WtStartLow OR #s130_WtPressProbesUp_T1) AND NOT #sStWtResetRel AND NOT #s140_WtStartLow_T1;
   IF #s140_WtStartLow THEN #qStateNo := 140; END_IF;
END_REGION

REGION Network 51: Actions for STATE Num:140 WtStartLow - qHiPotTestOver
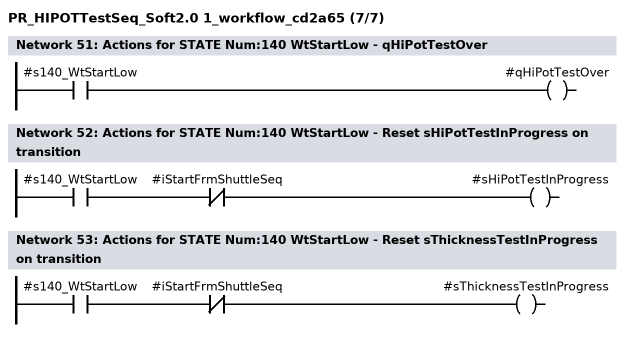
   RUNG wire#powerrail
      Contact( #s140_WtStartLow )
      Coil( #qHiPotTestOver )
   END_RUNG
   // the same network as SCL:
   #qHiPotTestOver := #s140_WtStartLow;
END_REGION

REGION Network 52: Actions for STATE Num:140 WtStartLow - Reset sHiPotTestInProgress on transition
   RUNG wire#powerrail
      Contact( #s140_WtStartLow )
      I_Contact( #iStartFrmShuttleSeq )
      Coil( #sHiPotTestInProgress )
   END_RUNG
   // the same network as SCL:
   #sHiPotTestInProgress := #s140_WtStartLow AND NOT #iStartFrmShuttleSeq;
END_REGION

REGION Network 53: Actions for STATE Num:140 WtStartLow - Reset sThicknessTestInProgress on transition
   RUNG wire#powerrail
      Contact( #s140_WtStartLow )
      I_Contact( #iStartFrmShuttleSeq )
      Coil( #sThicknessTestInProgress )
   END_RUNG
   // the same network as SCL:
   #sThicknessTestInProgress := #s140_WtStartLow AND NOT #iStartFrmShuttleSeq;
END_REGION
END_FUNCTION_BLOCK
